ADAPTER buttons (* Adapter Interface *)
  (* Standard: 61499-1 *)
  (* Version 0.0, 10/27/2026, lizar, Schneider Electric *)
  PACKAGE Main;
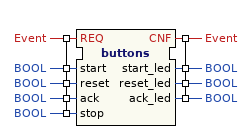
  EVENT_INPUT
    REQ WITH start, reset, ack, stop; (* Request from Socket *)
  END_EVENT
  EVENT_OUTPUT
    CNF WITH start_led, reset_led, ack_led; (* Confirmation from Plug *)
  END_EVENT
  VAR_INPUT
    start : BOOL; (* Request Data from Socket *)
    reset : BOOL; (* Response Data from Socket *)
    ack : BOOL; (* Response Data from Socket *)
    stop : BOOL; (* Response Data from Socket *)
  END_VAR
  VAR_OUTPUT
    start_led : BOOL; (* Confirmation Data from Plug *)
    reset_led : BOOL; (* Indication Data from Plug *)
    ack_led : BOOL; (* Indication Data from Plug *)
  END_VAR
  SERVICE SOCKET/PLUG
    SEQUENCE request_confirm
      SOCKET.REQ(start) -> PLUG.REQ(start);
      PLUG.CNF(start_led) -> SOCKET.CNF(start_led);
    END_SEQUENCE
    SEQUENCE indication_response
      PLUG.IND(reset_led) -> SOCKET.IND(reset_led);
      SOCKET.RSP(reset) -> PLUG.RSP(reset);
    END_SEQUENCE
  END_SERVICE
END_ADAPTER
